// Generated by voz_llm_plc_agent
// Target: Siemens TIA Portal V18 - SCL external source
// Review and compile before any download to physical hardware.

FUNCTION_BLOCK "PLC_PRG"
{ S7_Optimized_Access := 'TRUE' }
VERSION : 0.1
VAR_INPUT
   I_Start : Bool := FALSE;
   I_Emergency : Bool := FALSE;
END_VAR
VAR_OUTPUT
   Q_Motor_Enable : Bool := FALSE;
END_VAR
VAR
   T_DelayStart {InstructionName := 'TON_TIME'; LibVersion := '1.0'} : TON_TIME;
END_VAR
BEGIN
(* Arranque retardado del motor *)
#T_DelayStart(IN := #I_Start AND NOT FALSE AND NOT #I_Emergency, PT := T#3s);
#Q_Motor_Enable := #T_DelayStart.Q AND NOT FALSE AND NOT #I_Emergency;
(* Bloqueo: #I_Emergency fuerza a FALSE #Q_Motor_Enable de inmediato *)
IF #I_Emergency THEN
    #Q_Motor_Enable := FALSE;
END_IF;
END_FUNCTION_BLOCK

DATA_BLOCK "DB_PLC_PRG"
{ S7_Optimized_Access := 'TRUE' }
VERSION : 0.1
NON_RETAIN
"PLC_PRG"
BEGIN
END_DATA_BLOCK

ORGANIZATION_BLOCK "Main"
{ S7_Optimized_Access := 'TRUE' }
VERSION : 0.1
BEGIN
   "DB_PLC_PRG"(
      I_Start := "I_Start",
      I_Emergency := "I_Emergency",
      Q_Motor_Enable => "Q_Motor_Enable"
   );
END_ORGANIZATION_BLOCK
